FUNCTION_BLOCK ShortHandshake
VAR_INPUT
	ixStrobIn : BOOL;
END_VAR
VAR_OUTPUT
	oxStrobe : BOOL;
END_VAR
VAR
END_VAR

END_FUNCTION_BLOCK

(* stored: Version 1.1.0.1, ProductVersion 3.1.4024.12
   POU ShortHandshake: Id {ef228cbb-7e88-4e15-b0df-5963977c46cc}, SpecialFunc None *)
